ABB RobotStudio station: 260913Study1_0914_含Path_20.rsstn

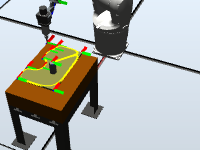
Station 260913Study1 (saved by RobotStudio 6.8.8148.134)
Controller 260913System1
  mechanical unit ROB_1: IRB1200_5_90_STD_02, 6 joints, base frame (0, 0, 0) mm
Layout (positions relative to the parent item):
  - IRB1200_5_90_STD_02 [mechanism, from Robots\IRB1200_5_90_STD_02.rslib] at (0, 0, 0) mm; joint values [-0.3705, 0.0008, 0.5103, 0.5015, 0.4822, -0.7492] (rad or m)
  - Curve_thing [part, from Training Objects\Curve_Thing.rslib] at (552.96, -150, 308) mm
  - table_and_fixture_140 [part, from Training Objects\propeller_table.rslib] at (527.96, -175, 0) mm
  - MyTool [mechanism, from Training Objects\myTool.rslib] at (436.63, -150, 598.53) mm, rotated rx 180 ry 38 rz 180 deg
Attachment: MyTool is attached to IRB1200_5_90_STD_02 / Link6
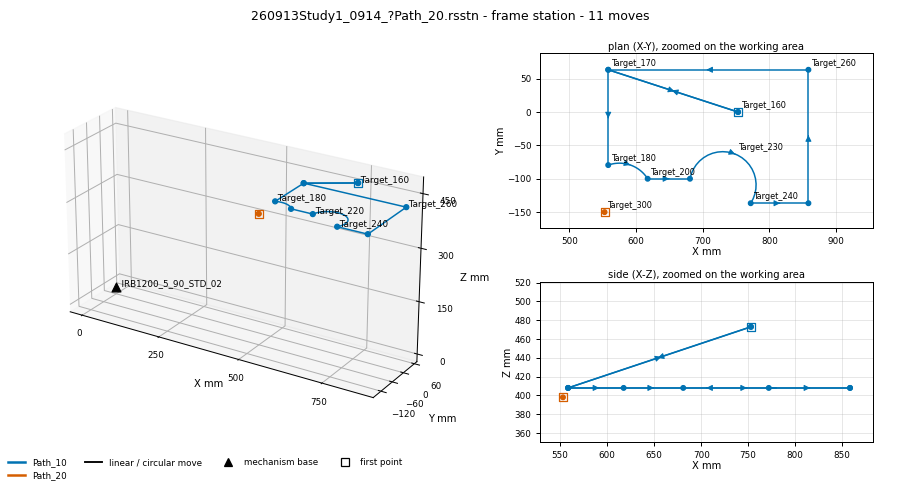
[picture p0: tool path of 260913Study1_0914_含Path_20.rsstn in frame station, 11 of 11 moves have a stored position in this frame; points joined in program order, loops and branches not executed]
Targets, tools, work objects and paths stored in the station, written as RAPID:
! task T_ROB1
MODULE CalibData
  PERS tooldata MyTool:=[TRUE,[[31.792631019,0,229.638935148],[0.945518576,0,0.325568154,0]],[1,[0,0,1],[1,0,0,0],0,0,0]];
ENDMODULE

! task T_ROB1
MODULE Module1
  CONST robtarget Target_160:=[[752.961021712,0,473.000001678],[-0.00000002,0,1,0],[0,-1,0,0],[9E+09,9E+09,9E+09,9E+09,9E+09,9E+09]];
  CONST robtarget Target_170:=[[558.409,63.326,408],[0,0,1,0],[0,-1,0,0],[9E+09,9E+09,9E+09,9E+09,9E+09,9E+09]];
  CONST robtarget Target_180:=[[558.409,-79.547,408],[0,0,1,0],[-1,0,-1,0],[9E+09,9E+09,9E+09,9E+09,9E+09,9E+09]];
  CONST robtarget Target_190:=[[591.551,-79.397,408],[0,0,1,0],[-1,0,-1,0],[9E+09,9E+09,9E+09,9E+09,9E+09,9E+09]];
  CONST robtarget Target_200:=[[617.506,-100.006,408],[0,0,1,0],[-1,0,-1,0],[9E+09,9E+09,9E+09,9E+09,9E+09,9E+09]];
  CONST robtarget Target_210:=[[752.961,0,473],[0,0,1,0],[0,0,0,0],[9E+09,9E+09,9E+09,9E+09,9E+09,9E+09]];
  CONST robtarget Target_220:=[[680.926,-100.006,408],[0,0,1,0],[0,0,0,0],[9E+09,9E+09,9E+09,9E+09,9E+09,9E+09]];
  CONST robtarget Target_230:=[[748.721,-63.019,408],[0,0,1,0],[0,0,0,0],[9E+09,9E+09,9E+09,9E+09,9E+09,9E+09]];
  CONST robtarget Target_240:=[[771.941,-136.674,408],[0,0,1,0],[0,0,0,0],[9E+09,9E+09,9E+09,9E+09,9E+09,9E+09]];
  CONST robtarget Target_250:=[[858.409,-136.674,408],[0,0,1,0],[0,0,0,0],[9E+09,9E+09,9E+09,9E+09,9E+09,9E+09]];
  CONST robtarget Target_260:=[[858.409,63.326,408],[0,0,1,0],[0,0,0,0],[9E+09,9E+09,9E+09,9E+09,9E+09,9E+09]];
  CONST robtarget Target_270:=[[558.409,63.326,408],[0,0,1,0],[0,0,0,0],[9E+09,9E+09,9E+09,9E+09,9E+09,9E+09]];
  CONST robtarget Target_280:=[[752.961,0,473],[0,0,1,0],[0,0,0,0],[9E+09,9E+09,9E+09,9E+09,9E+09,9E+09]];
  CONST robtarget Target_290:=[[552.961,-150,398],[-0.00000002,0,1,0],[0,0,0,0],[9E+09,9E+09,9E+09,9E+09,9E+09,9E+09]];
  CONST robtarget Target_300:=[[552.961,-150,398],[-0.00000002,0,1,0],[0,0,0,0],[9E+09,9E+09,9E+09,9E+09,9E+09,9E+09]];
  PROC Path_10()
    MoveJ Target_160,v50,z100,MyTool\WObj:=wobj0;
    MoveL Target_170,v50,z100,MyTool\WObj:=wobj0;
    MoveL Target_180,v50,z100,MyTool\WObj:=wobj0;
    MoveC Target_190,Target_200,v50,z100,MyTool\WObj:=wobj0;
    MoveL Target_220,v50,z100,MyTool\WObj:=wobj0;
    MoveC Target_230,Target_240,v50,z100,MyTool\WObj:=wobj0;
    MoveL Target_250,v50,z100,MyTool\WObj:=wobj0;
    MoveL Target_260,v50,z100,MyTool\WObj:=wobj0;
    MoveL Target_270,v50,z100,MyTool\WObj:=wobj0;
    MoveL Target_280,v50,z100,MyTool\WObj:=wobj0;
  ENDPROC
  PROC Path_20()
    MoveL Target_300,v50,z100,MyTool\WObj:=wobj0;
  ENDPROC
ENDMODULE

